--- program cerlatderch (robot Fanuc LR Mate 200iD/7L) ---
  Suave(1)
  Establecer velocidad (1000.0 mm/s)
  Est. Ref.: RobotiQ 2F-140 Gripper (Mechanism) Base
  Est. herr: Tool 1
  Mostrar Tool 1
  MoveJ 1 to (255.53, 172.79, 254.67) mm, rotated rx 167 ry -29.36 rz -83.53 deg; joints [62.819, 42.709, -13.957, -31.792, -82.544, 126.287]
  MoveL 2 to (255.53, 172.79, 254.67) mm, rotated rx 167 ry -29.36 rz -83.53 deg; joints [62.819, 42.709, -13.957, -31.792, -82.544, 126.287]
  MoveL 3 to (235.92, 172.79, 156.61) mm, rotated rx 167 ry -29.36 rz -83.53 deg; joints [63.476, 48.891, -22.926, -32.864, -74.628, 130.64]
  MoveL 4 to (235.92, 172.79, 156.61) mm, rotated rx 167 ry -29.36 rz -83.53 deg; joints [63.476, 48.891, -22.926, -32.864, -74.628, 130.64]
  Establecer velocidad (50.0 mm/s)
  MoveL 5 to (245.19, 173.88, 156.61) mm, rotated rx 167 ry -29.36 rz -83.53 deg; joints [63.097, 47.784, -23.838, -32.935, -74.051, 131.456]
  MoveL 6 to (254.51, 174, 156.61) mm, rotated rx 167 ry -29.36 rz -83.53 deg; joints [62.774, 46.641, -24.767, -33.021, -73.432, 132.241]
  MoveL 7 to (263.84, 173.92, 156.61) mm, rotated rx 167 ry -29.36 rz -83.53 deg; joints [62.457, 45.515, -25.67, -33.109, -72.832, 133.007]
  MoveL 8 to (273.13, 173.41, 156.77) mm, rotated rx 167 ry -29.36 rz -83.53 deg; joints [62.163, 44.386, -26.542, -33.199, -72.246, 133.739]
  MoveL 9 to (282.79, 172.36, 157.79) mm, rotated rx 167 ry -29.36 rz -83.53 deg; joints [61.885, 43.161, -27.346, -33.284, -71.709, 134.42]
  MoveL 10 to (292.21, 170.83, 159.74) mm, rotated rx 167 ry -29.36 rz -83.53 deg; joints [61.643, 41.908, -28.02, -33.355, -71.264, 134.999]
  MoveL 11 to (301.4, 168.84, 162.6) mm, rotated rx 167 ry -29.36 rz -83.53 deg; joints [61.436, 40.621, -28.563, -33.411, -70.911, 135.476]
  MoveL 12 to (310.49, 166.4, 165.63) mm, rotated rx 167 ry -29.36 rz -83.53 deg; joints [61.259, 39.322, -29.065, -33.468, -70.577, 135.906]
  MoveL 13 to (319.81, 164.14, 167.77) mm, rotated rx 167 ry -29.36 rz -83.53 deg; joints [61.056, 38.072, -29.642, -33.535, -70.194, 136.401]
  MoveL 14 to (329.36, 162.38, 169) mm, rotated rx 167 ry -29.36 rz -83.53 deg; joints [60.801, 36.892, -30.285, -33.604, -69.78, 136.975]
  MoveL 15 to (339.84, 161.1, 169.31) mm, rotated rx 167 ry -29.36 rz -83.53 deg; joints [60.468, 35.712, -31.049, -33.681, -69.303, 137.681]
  MoveL 16 to (350.39, 160.46, 169.31) mm, rotated rx 167 ry -29.36 rz -83.53 deg; joints [60.074, 34.597, -31.799, -33.741, -68.866, 138.426]
  MoveL 17 to (360.96, 160.39, 169.31) mm, rotated rx 167 ry -29.36 rz -83.53 deg; joints [59.626, 33.529, -32.502, -33.778, -68.492, 139.185]
  MoveL 18 to (371.53, 160.39, 169.31) mm, rotated rx 167 ry -29.36 rz -83.53 deg; joints [59.16, 32.48, -33.179, -33.805, -68.148, 139.94]
  MoveL 19 to (382.1, 160.39, 169.31) mm, rotated rx 167 ry -29.36 rz -83.53 deg; joints [58.681, 31.444, -33.831, -33.821, -67.828, 140.689]
  MoveL 20 to (408.52, 160.39, 169.31) mm, rotated rx 167 ry -29.36 rz -83.53 deg; joints [57.423, 28.911, -35.364, -33.817, -67.131, 142.544]
  MoveL 21 to (413.03, 160.03, 169.31) mm, rotated rx 167 ry -29.36 rz -83.53 deg; joints [57.227, 28.464, -35.624, -33.821, -67.004, 142.845]
  MoveL 22 to (417.64, 158.65, 169.31) mm, rotated rx 167 ry -29.36 rz -83.53 deg; joints [57.103, 27.947, -35.922, -33.855, -66.812, 143.116]
  MoveL 23 to (422.01, 156.15, 169.31) mm, rotated rx 167 ry -29.36 rz -83.53 deg; joints [57.077, 27.387, -36.239, -33.923, -66.56, 143.328]
  MoveL 24 to (425.74, 152.66, 169.31) mm, rotated rx 167 ry -29.36 rz -83.53 deg; joints [57.162, 26.828, -36.552, -34.025, -66.262, 143.456]
  MoveL 25 to (428.54, 148.44, 169.31) mm, rotated rx 167 ry -29.36 rz -83.53 deg; joints [57.356, 26.314, -36.835, -34.154, -65.941, 143.489]
  MoveL 26 to (430.23, 143.87, 169.31) mm, rotated rx 167 ry -29.36 rz -83.53 deg; joints [57.636, 25.883, -37.068, -34.299, -65.622, 143.43]
  MoveL 27 to (430.87, 139.33, 169.31) mm, rotated rx 167 ry -29.36 rz -83.53 deg; joints [57.973, 25.556, -37.244, -34.446, -65.326, 143.295]
  MoveL 28 to (430.88, 134.93, 169.31) mm, rotated rx 167 ry -29.36 rz -83.53 deg; joints [58.333, 25.298, -37.381, -34.591, -65.05, 143.121]
  MoveL 29 to (430.86, 130.52, 169.31) mm, rotated rx 167 ry -29.36 rz -83.53 deg; joints [58.698, 25.045, -37.514, -34.737, -64.776, 142.942]
  MoveL 30 to (430.2, 125.97, 169.31) mm, rotated rx 167 ry -29.36 rz -83.53 deg; joints [59.109, 24.848, -37.618, -34.889, -64.505, 142.711]
  MoveL 31 to (428.47, 121.41, 169.31) mm, rotated rx 167 ry -29.36 rz -83.53 deg; joints [59.577, 24.755, -37.666, -35.042, -64.253, 142.405]
  MoveL 32 to (425.65, 117.21, 169.31) mm, rotated rx 167 ry -29.36 rz -83.53 deg; joints [60.069, 24.791, -37.647, -35.183, -64.045, 142.039]
  MoveL 33 to (421.9, 113.74, 169.31) mm, rotated rx 167 ry -29.36 rz -83.53 deg; joints [60.543, 24.962, -37.558, -35.297, -63.901, 141.64]
  MoveL 34 to (417.52, 111.28, 169.31) mm, rotated rx 167 ry -29.36 rz -83.53 deg; joints [60.959, 25.251, -37.405, -35.375, -63.834, 141.242]
  MoveL 35 to (412.24, 109.81, 169.31) mm, rotated rx 167 ry -29.36 rz -83.53 deg; joints [61.327, 25.684, -37.175, -35.415, -63.852, 140.827]
  MoveL 36 to (407.14, 109.59, 169.31) mm, rotated rx 167 ry -29.36 rz -83.53 deg; joints [61.58, 26.169, -36.913, -35.413, -63.949, 140.475]
  MoveL 37 to (402.11, 109.59, 169.31) mm, rotated rx 167 ry -29.36 rz -83.53 deg; joints [61.806, 26.66, -36.644, -35.4, -64.063, 140.137]
  MoveL 38 to (397.07, 109.59, 169.31) mm, rotated rx 167 ry -29.36 rz -83.53 deg; joints [62.03, 27.154, -36.37, -35.385, -64.183, 139.798]
  MoveL 39 to (392.04, 109.59, 169.31) mm, rotated rx 167 ry -29.36 rz -83.53 deg; joints [62.25, 27.65, -36.091, -35.367, -64.308, 139.458]
  MoveL 40 to (387.01, 109.59, 169.31) mm, rotated rx 167 ry -29.36 rz -83.53 deg; joints [62.467, 28.147, -35.807, -35.347, -64.438, 139.117]
  MoveL 41 to (381.98, 109.59, 169.31) mm, rotated rx 167 ry -29.36 rz -83.53 deg; joints [62.681, 28.647, -35.517, -35.325, -64.573, 138.774]
  MoveL 42 to (370.35, 109.59, 169.31) mm, rotated rx 167 ry -29.36 rz -83.53 deg; joints [63.163, 29.81, -34.83, -35.263, -64.906, 137.979]
  MoveL 43 to (358.72, 109.59, 169.31) mm, rotated rx 167 ry -29.36 rz -83.53 deg; joints [63.63, 30.986, -34.115, -35.19, -65.268, 137.178]
  MoveL 44 to (347.1, 109.76, 169.31) mm, rotated rx 167 ry -29.36 rz -83.53 deg; joints [64.069, 32.184, -33.366, -35.101, -65.671, 136.376]
  MoveL 45 to (335.47, 109.5, 169.3) mm, rotated rx 167 ry -29.36 rz -83.53 deg; joints [64.527, 33.378, -32.602, -35.013, -66.075, 135.551]
  MoveL 46 to (325.71, 108.73, 168.64) mm, rotated rx 167 ry -29.36 rz -83.53 deg; joints [64.943, 34.406, -32.028, -34.963, -66.344, 134.876]
  MoveL 47 to (316.17, 107.5, 167.04) mm, rotated rx 167 ry -29.36 rz -83.53 deg; joints [65.376, 35.455, -31.568, -34.945, -66.51, 134.259]
  MoveL 48 to (306.86, 105.82, 164.53) mm, rotated rx 167 ry -29.36 rz -83.53 deg; joints [65.826, 36.522, -31.218, -34.955, -66.577, 133.698]
  MoveL 49 to (297.74, 103.7, 161.34) mm, rotated rx 167 ry -29.36 rz -83.53 deg; joints [66.291, 37.598, -30.947, -34.987, -66.571, 133.172]
  MoveL 50 to (288.57, 101.1, 158.87) mm, rotated rx 167 ry -29.36 rz -83.53 deg; joints [66.786, 38.625, -30.584, -34.999, -66.625, 132.566]
  MoveL 51 to (279.32, 97.99, 157.31) mm, rotated rx 167 ry -29.36 rz -83.53 deg; joints [67.309, 39.597, -30.108, -34.986, -66.755, 131.867]
  MoveL 52 to (269.16, 95.14, 156.63) mm, rotated rx 167 ry -29.36 rz -83.53 deg; joints [67.83, 40.652, -29.429, -34.921, -67.053, 131.04]
  MoveL 53 to (258.73, 93.27, 156.61) mm, rotated rx 167 ry -29.36 rz -83.53 deg; joints [68.276, 41.767, -28.59, -34.803, -67.518, 130.173]
  MoveL 54 to (248.13, 92.41, 156.61) mm, rotated rx 167 ry -29.36 rz -83.53 deg; joints [68.643, 42.973, -27.665, -34.652, -68.094, 129.318]
  MoveL 55 to (237.5, 92.57, 156.61) mm, rotated rx 167 ry -29.36 rz -83.53 deg; joints [68.927, 44.261, -26.662, -34.475, -68.777, 128.482]
  MoveL 56 to (226.98, 93.76, 156.67) mm, rotated rx 167 ry -29.36 rz -83.53 deg; joints [69.129, 45.614, -25.583, -34.275, -69.565, 127.669]
  MoveL 57 to (220.53, 95, 156.94) mm, rotated rx 167 ry -29.36 rz -83.53 deg; joints [69.214, 46.476, -24.851, -34.137, -70.127, 127.164]
  MoveL 58 to (214.18, 96.62, 157.45) mm, rotated rx 167 ry -29.36 rz -83.53 deg; joints [69.269, 47.348, -24.072, -33.99, -70.745, 126.656]
  MoveL 59 to (207.94, 98.62, 158.18) mm, rotated rx 167 ry -29.36 rz -83.53 deg; joints [69.294, 48.235, -23.243, -33.835, -71.42, 126.147]
  MoveL 60 to (202.03, 101.35, 159.07) mm, rotated rx 167 ry -29.36 rz -83.53 deg; joints [69.26, 49.127, -22.379, -33.672, -72.155, 125.67]
  MoveL 61 to (196.78, 105.2, 160.04) mm, rotated rx 167 ry -29.36 rz -83.53 deg; joints [69.133, 50.007, -21.509, -33.504, -72.945, 125.267]
  MoveL 62 to (192.41, 110, 160.98) mm, rotated rx 167 ry -29.36 rz -83.53 deg; joints [68.923, 50.84, -20.677, -33.341, -73.747, 124.96]
  MoveL 63 to (189.05, 115.61, 161.78) mm, rotated rx 167 ry -29.36 rz -83.53 deg; joints [68.635, 51.604, -19.92, -33.187, -74.529, 124.763]
  MoveL 64 to (186.87, 121.77, 162.34) mm, rotated rx 167 ry -29.36 rz -83.53 deg; joints [68.284, 52.257, -19.287, -33.05, -75.24, 124.692]
  MoveL 65 to (186.12, 126.11, 162.54) mm, rotated rx 167 ry -29.36 rz -83.53 deg; joints [68.018, 52.62, -18.948, -32.97, -75.661, 124.719]
  MoveL 66 to (185.93, 130.52, 162.58) mm, rotated rx 167 ry -29.36 rz -83.53 deg; joints [67.733, 52.914, -18.69, -32.9, -76.024, 124.807]
  MoveL 67 to (186.01, 134.94, 162.56) mm, rotated rx 167 ry -29.36 rz -83.53 deg; joints [67.443, 53.178, -18.465, -32.834, -76.362, 124.92]
  MoveL 68 to (186.83, 139.23, 162.35) mm, rotated rx 167 ry -29.36 rz -83.53 deg; joints [67.141, 53.335, -18.361, -32.783, -76.605, 125.109]
  MoveL 69 to (189.27, 144.53, 161.73) mm, rotated rx 167 ry -29.36 rz -83.53 deg; joints [66.73, 53.332, -18.45, -32.742, -76.741, 125.496]
  MoveL 70 to (192.92, 149.04, 160.87) mm, rotated rx 167 ry -29.36 rz -83.53 deg; joints [66.335, 53.113, -18.76, -32.73, -76.683, 125.992]
  MoveL 71 to (196.97, 153.16, 160.01) mm, rotated rx 167 ry -29.36 rz -83.53 deg; joints [65.952, 52.817, -19.134, -32.727, -76.564, 126.513]
  MoveL 72 to (203.59, 158.73, 158.82) mm, rotated rx 167 ry -29.36 rz -83.53 deg; joints [65.398, 52.27, -19.77, -32.731, -76.311, 127.319]
  MoveL 73 to (210.87, 163.56, 157.81) mm, rotated rx 167 ry -29.36 rz -83.53 deg; joints [64.867, 51.598, -20.485, -32.747, -75.979, 128.149]
  MoveL 74 to (218.67, 167.53, 157.07) mm, rotated rx 167 ry -29.36 rz -83.53 deg; joints [64.37, 50.814, -21.254, -32.774, -75.585, 128.981]
  MoveL 75 to (226.86, 170.59, 156.67) mm, rotated rx 167 ry -29.36 rz -83.53 deg; joints [63.913, 49.93, -22.054, -32.812, -75.142, 129.798]
  Establecer velocidad (1000.0 mm/s)
  MoveL 76 to (226.86, 170.59, 156.67) mm, rotated rx 167 ry -29.36 rz -83.53 deg; joints [63.913, 49.93, -22.054, -32.812, -75.142, 129.798]
  MoveL 77 to (246.47, 170.59, 254.73) mm, rotated rx 167 ry -29.36 rz -83.53 deg; joints [63.272, 43.813, -13.15, -31.797, -82.998, 125.482]
  Establecer velocidad (1000.0 mm/s)
  MoveL 78 to (401.83, 160.52, 306.49) mm, rotated rx 167 ry -29.36 rz -83.53 deg; joints [57.739, 22.896, -18.143, -31.275, -81.532, 132.699]
  MoveL 79 to (382.22, 160.52, 208.44) mm, rotated rx 167 ry -29.36 rz -83.53 deg; joints [58.665, 29.141, -29.231, -32.884, -71.679, 138.006]
  MoveL 80 to (382.22, 160.52, 208.44) mm, rotated rx 167 ry -29.36 rz -83.53 deg; joints [58.665, 29.141, -29.231, -32.884, -71.679, 138.006]
  Establecer velocidad (50.0 mm/s)
  MoveL 81 to (398.1, 159.77, 208.44) mm, rotated rx 167 ry -29.36 rz -83.53 deg; joints [57.977, 27.495, -30.13, -32.875, -71.248, 139.05]
  MoveL 82 to (413.85, 157.57, 208.44) mm, rotated rx 167 ry -29.36 rz -83.53 deg; joints [57.377, 25.796, -31.013, -32.884, -70.787, 140.016]
  MoveL 83 to (418.98, 156.18, 208.44) mm, rotated rx 167 ry -29.36 rz -83.53 deg; joints [57.228, 25.206, -31.31, -32.901, -70.607, 140.3]
  MoveL 84 to (423.65, 153.71, 208.44) mm, rotated rx 167 ry -29.36 rz -83.53 deg; joints [57.186, 24.593, -31.611, -32.947, -70.373, 140.506]
  MoveL 85 to (427.7, 150.29, 208.44) mm, rotated rx 167 ry -29.36 rz -83.53 deg; joints [57.25, 23.982, -31.906, -33.022, -70.097, 140.627]
  MoveL 86 to (430.9, 146.07, 208.44) mm, rotated rx 167 ry -29.36 rz -83.53 deg; joints [57.424, 23.406, -32.178, -33.124, -69.788, 140.654]
  MoveL 87 to (432.92, 141.18, 208.44) mm, rotated rx 167 ry -29.36 rz -83.53 deg; joints [57.717, 22.905, -32.409, -33.25, -69.459, 140.568]
  MoveL 88 to (433.51, 135.92, 208.44) mm, rotated rx 167 ry -29.36 rz -83.53 deg; joints [58.117, 22.524, -32.583, -33.395, -69.128, 140.369]
  MoveL 89 to (433.26, 130.66, 208.44) mm, rotated rx 167 ry -29.36 rz -83.53 deg; joints [58.565, 22.229, -32.715, -33.544, -68.81, 140.11]
  MoveL 90 to (431.75, 125.64, 208.44) mm, rotated rx 167 ry -29.36 rz -83.53 deg; joints [59.059, 22.078, -32.783, -33.69, -68.524, 139.778]
  MoveL 91 to (428.97, 121.16, 208.44) mm, rotated rx 167 ry -29.36 rz -83.53 deg; joints [59.573, 22.09, -32.777, -33.825, -68.288, 139.389]
  MoveL 92 to (425.29, 117.41, 208.44) mm, rotated rx 167 ry -29.36 rz -83.53 deg; joints [60.069, 22.241, -32.71, -33.94, -68.111, 138.975]
  MoveL 93 to (421.02, 114.59, 208.44) mm, rotated rx 167 ry -29.36 rz -83.53 deg; joints [60.513, 22.508, -32.59, -34.027, -68.002, 138.569]
  MoveL 94 to (416.24, 112.78, 208.44) mm, rotated rx 167 ry -29.36 rz -83.53 deg; joints [60.891, 22.888, -32.417, -34.085, -67.967, 138.179]
  MoveL 95 to (411.24, 111.87, 208.44) mm, rotated rx 167 ry -29.36 rz -83.53 deg; joints [61.2, 23.343, -32.206, -34.115, -67.995, 137.819]
  MoveL 96 to (406.21, 111.14, 208.44) mm, rotated rx 167 ry -29.36 rz -83.53 deg; joints [61.491, 23.815, -31.985, -34.137, -68.04, 137.464]
  MoveL 97 to (393.32, 109.92, 208.44) mm, rotated rx 167 ry -29.36 rz -83.53 deg; joints [62.167, 25.068, -31.378, -34.164, -68.22, 136.585]
  MoveL 98 to (380.38, 109.57, 208.44) mm, rotated rx 167 ry -29.36 rz -83.53 deg; joints [62.749, 26.389, -30.71, -34.151, -68.492, 135.737]
  MoveL 99 to (368.61, 109.92, 208.44) mm, rotated rx 167 ry -29.36 rz -83.53 deg; joints [63.207, 27.639, -30.053, -34.111, -68.815, 134.99]
  MoveL 100 to (356.97, 111.21, 208.44) mm, rotated rx 167 ry -29.36 rz -83.53 deg; joints [63.57, 28.939, -29.343, -34.038, -69.225, 134.285]
  MoveL 101 to (345.55, 113.37, 208.44) mm, rotated rx 167 ry -29.36 rz -83.53 deg; joints [63.844, 30.275, -28.588, -33.939, -69.717, 133.622]
  MoveL 102 to (333.92, 113.25, 208.44) mm, rotated rx 167 ry -29.36 rz -83.53 deg; joints [64.293, 31.528, -27.855, -33.881, -70.105, 132.837]
  MoveL 103 to (322.29, 113.18, 208.44) mm, rotated rx 167 ry -29.36 rz -83.53 deg; joints [64.724, 32.803, -27.087, -33.814, -70.53, 132.045]
  MoveL 104 to (318.84, 113.27, 208.44) mm, rotated rx 167 ry -29.36 rz -83.53 deg; joints [64.842, 33.192, -26.849, -33.79, -70.669, 131.812]
  MoveL 105 to (315.38, 113.44, 208.44) mm, rotated rx 167 ry -29.36 rz -83.53 deg; joints [64.952, 33.586, -26.605, -33.763, -70.818, 131.582]
  MoveL 106 to (311.94, 113.73, 208.44) mm, rotated rx 167 ry -29.36 rz -83.53 deg; joints [65.051, 33.988, -26.353, -33.733, -70.977, 131.356]
  MoveL 107 to (308.53, 114.29, 208.44) mm, rotated rx 167 ry -29.36 rz -83.53 deg; joints [65.128, 34.401, -26.093, -33.698, -71.156, 131.142]
  MoveL 108 to (305.51, 115.94, 208.44) mm, rotated rx 167 ry -29.36 rz -83.53 deg; joints [65.11, 34.829, -25.821, -33.644, -71.391, 130.998]
  MoveL 109 to (303.55, 118.04, 208.44) mm, rotated rx 167 ry -29.36 rz -83.53 deg; joints [65.021, 35.163, -25.606, -33.588, -71.614, 130.943]
  MoveL 110 to (302.26, 120.61, 208.44) mm, rotated rx 167 ry -29.36 rz -83.53 deg; joints [64.874, 35.447, -25.423, -33.528, -71.84, 130.952]
  MoveL 111 to (301.89, 123.45, 208.44) mm, rotated rx 167 ry -29.36 rz -83.53 deg; joints [64.677, 35.642, -25.297, -33.469, -72.044, 131.035]
  MoveL 112 to (302.49, 126.27, 208.44) mm, rotated rx 167 ry -29.36 rz -83.53 deg; joints [64.448, 35.726, -25.242, -33.417, -72.204, 131.185]
  MoveL 113 to (303.41, 129.02, 208.44) mm, rotated rx 167 ry -29.36 rz -83.53 deg; joints [64.213, 35.772, -25.213, -33.368, -72.345, 131.354]
  MoveL 114 to (304.36, 131.76, 208.44) mm, rotated rx 167 ry -29.36 rz -83.53 deg; joints [63.978, 35.816, -25.184, -33.32, -72.486, 131.524]
  MoveL 115 to (304.62, 133.96, 208.44) mm, rotated rx 167 ry -29.36 rz -83.53 deg; joints [63.808, 35.909, -25.123, -33.277, -72.621, 131.624]
  MoveL 116 to (303.96, 136.18, 208.44) mm, rotated rx 167 ry -29.36 rz -83.53 deg; joints [63.669, 36.109, -24.993, -33.229, -72.799, 131.659]
  MoveL 117 to (303.31, 138.41, 208.44) mm, rotated rx 167 ry -29.36 rz -83.53 deg; joints [63.531, 36.308, -24.862, -33.181, -72.978, 131.694]
  MoveL 118 to (302.68, 140.64, 208.44) mm, rotated rx 167 ry -29.36 rz -83.53 deg; joints [63.392, 36.507, -24.73, -33.133, -73.157, 131.729]
  MoveL 119 to (302.1, 142.88, 208.44) mm, rotated rx 167 ry -29.36 rz -83.53 deg; joints [63.251, 36.703, -24.601, -33.085, -73.335, 131.767]
  MoveL 120 to (302.05, 146.74, 208.44) mm, rotated rx 167 ry -29.36 rz -83.53 deg; joints [62.975, 36.931, -24.449, -33.008, -73.599, 131.9]
  MoveL 121 to (303.35, 150.38, 208.44) mm, rotated rx 167 ry -29.36 rz -83.53 deg; joints [62.667, 36.996, -24.406, -32.943, -73.788, 132.121]
  MoveL 122 to (305.63, 153.5, 208.44) mm, rotated rx 167 ry -29.36 rz -83.53 deg; joints [62.359, 36.922, -24.455, -32.892, -73.899, 132.394]
  MoveL 123 to (308.22, 155.56, 208.44) mm, rotated rx 167 ry -29.36 rz -83.53 deg; joints [62.114, 36.75, -24.569, -32.862, -73.924, 132.653]
  MoveL 124 to (311.4, 156.56, 208.44) mm, rotated rx 167 ry -29.36 rz -83.53 deg; joints [61.923, 36.452, -24.767, -32.855, -73.852, 132.917]
  MoveL 125 to (314.73, 157, 208.44) mm, rotated rx 167 ry -29.36 rz -83.53 deg; joints [61.763, 36.105, -24.995, -32.859, -73.739, 133.172]
  MoveL 126 to (318.08, 157.27, 208.44) mm, rotated rx 167 ry -29.36 rz -83.53 deg; joints [61.615, 35.747, -25.229, -32.866, -73.616, 133.422]
  MoveL 127 to (321.43, 157.41, 208.44) mm, rotated rx 167 ry -29.36 rz -83.53 deg; joints [61.474, 35.383, -25.465, -32.876, -73.487, 133.667]
  MoveL 128 to (324.78, 157.45, 208.44) mm, rotated rx 167 ry -29.36 rz -83.53 deg; joints [61.34, 35.016, -25.701, -32.886, -73.354, 133.907]
  MoveL 129 to (328.13, 157.42, 208.44) mm, rotated rx 167 ry -29.36 rz -83.53 deg; joints [61.209, 34.647, -25.937, -32.897, -73.22, 134.144]
  MoveL 130 to (335.01, 157.24, 208.44) mm, rotated rx 167 ry -29.36 rz -83.53 deg; joints [60.946, 33.887, -26.417, -32.921, -72.945, 134.624]
  MoveL 131 to (341.89, 157.02, 208.44) mm, rotated rx 167 ry -29.36 rz -83.53 deg; joints [60.681, 33.133, -26.886, -32.942, -72.681, 135.099]
  MoveL 132 to (348.73, 157.41, 208.44) mm, rotated rx 167 ry -29.36 rz -83.53 deg; joints [60.368, 32.427, -27.317, -32.947, -72.47, 135.589]
  MoveL 133 to (355.61, 159.03, 208.44) mm, rotated rx 167 ry -29.36 rz -83.53 deg; joints [59.957, 31.799, -27.695, -32.919, -72.351, 136.126]
  MoveL 134 to (359.78, 159.91, 208.44) mm, rotated rx 167 ry -29.36 rz -83.53 deg; joints [59.712, 31.415, -27.923, -32.902, -72.277, 136.447]
  MoveL 135 to (363.08, 160.33, 208.44) mm, rotated rx 167 ry -29.36 rz -83.53 deg; joints [59.538, 31.096, -28.111, -32.894, -72.203, 136.69]
  MoveL 136 to (365.62, 160.48, 208.44) mm, rotated rx 167 ry -29.36 rz -83.53 deg; joints [59.414, 30.842, -28.26, -32.891, -72.137, 136.871]
  MoveL 137 to (367.82, 160.52, 208.44) mm, rotated rx 167 ry -29.36 rz -83.53 deg; joints [59.315, 30.617, -28.391, -32.891, -72.075, 137.023]
  MoveL 138 to (370.1, 160.52, 208.44) mm, rotated rx 167 ry -29.36 rz -83.53 deg; joints [59.213, 30.381, -28.527, -32.891, -72.009, 137.18]
  MoveL 139 to (372.32, 160.52, 208.44) mm, rotated rx 167 ry -29.36 rz -83.53 deg; joints [59.114, 30.153, -28.659, -32.89, -71.946, 137.332]
  MoveL 140 to (375.19, 160.52, 208.44) mm, rotated rx 167 ry -29.36 rz -83.53 deg; joints [58.985, 29.859, -28.827, -32.889, -71.866, 137.527]
  MoveL 141 to (378.62, 160.52, 208.44) mm, rotated rx 167 ry -29.36 rz -83.53 deg; joints [58.83, 29.508, -29.025, -32.887, -71.773, 137.761]
  MoveL 142 to (382.22, 160.52, 208.44) mm, rotated rx 167 ry -29.36 rz -83.53 deg; joints [58.665, 29.141, -29.231, -32.884, -71.679, 138.006]
  Establecer velocidad (1000.0 mm/s)
  MoveL 143 to (382.22, 160.52, 208.44) mm, rotated rx 167 ry -29.36 rz -83.53 deg; joints [58.665, 29.141, -29.231, -32.884, -71.679, 138.006]
  MoveL 144 to (401.83, 160.52, 306.49) mm, rotated rx 167 ry -29.36 rz -83.53 deg; joints [57.739, 22.896, -18.143, -31.275, -81.532, 132.699]

--- program ceraarribderch (robot Fanuc LR Mate 200iD/7L) ---
  Suave(1)
  Establecer velocidad (1000.0 mm/s)
  Est. Ref.: bote cera
  Est. herr: Tool 1
  Mostrar Tool 1
  MoveJ 1 to (349.44, 103.38, 195.99) mm, rotated rx 122.56 ry -24.48 rz -84.76 deg; joints [61.244, 18.633, -53.476, -104.529, -42.664, -159.742]
  MoveL 2 to (349.44, 103.38, 195.99) mm, rotated rx 122.56 ry -24.48 rz -84.76 deg; joints [61.244, 18.633, -53.476, -104.529, -42.664, -159.742]
  MoveL 3 to (329.83, 103.38, 97.93) mm, rotated rx 122.56 ry -24.48 rz -84.76 deg; joints [62.357, 32.195, -66.199, -117.758, -46.769, -142.563]
  MoveL 4 to (329.83, 103.38, 97.93) mm, rotated rx 122.56 ry -24.48 rz -84.76 deg; joints [62.357, 32.195, -66.199, -117.758, -46.769, -142.563]
  Establecer velocidad (50.0 mm/s)
  MoveL 5 to (328.15, 103.38, 97.77) mm, rotated rx 122.56 ry -24.48 rz -84.76 deg; joints [62.448, 32.321, -66.096, -117.772, -46.689, -142.664]
  MoveL 6 to (326.47, 103.38, 97.62) mm, rotated rx 122.56 ry -24.48 rz -84.76 deg; joints [62.539, 32.448, -65.992, -117.785, -46.608, -142.766]
  MoveL 7 to (322.21, 103.38, 97.19) mm, rotated rx 122.56 ry -24.48 rz -84.76 deg; joints [62.767, 32.775, -65.732, -117.817, -46.404, -143.023]
  MoveL 8 to (312.54, 103.38, 96.02) mm, rotated rx 122.56 ry -24.48 rz -84.76 deg; joints [63.273, 33.544, -65.159, -117.885, -45.95, -143.589]
  MoveL 9 to (290.7, 103.38, 92.42) mm, rotated rx 122.56 ry -24.48 rz -84.76 deg; joints [64.353, 35.413, -63.937, -118.011, -44.967, -144.799]
  MoveL 10 to (282.18, 103.38, 90.65) mm, rotated rx 122.56 ry -24.48 rz -84.76 deg; joints [64.752, 36.19, -63.484, -118.051, -44.599, -145.248]
  MoveL 11 to (277.43, 103.38, 89.57) mm, rotated rx 122.56 ry -24.48 rz -84.76 deg; joints [64.97, 36.634, -63.237, -118.07, -44.396, -145.494]
  MoveL 12 to (274.78, 103.38, 88.94) mm, rotated rx 122.56 ry -24.48 rz -84.76 deg; joints [65.09, 36.886, -63.101, -118.08, -44.284, -145.63]
  MoveL 13 to (273.09, 103.38, 88.53) mm, rotated rx 122.56 ry -24.48 rz -84.76 deg; joints [65.166, 37.048, -63.014, -118.086, -44.213, -145.715]
  MoveL 14 to (271.43, 103.38, 88.06) mm, rotated rx 122.56 ry -24.48 rz -84.76 deg; joints [65.24, 37.215, -62.937, -118.098, -44.147, -145.791]
  MoveL 15 to (269.69, 103.38, 86.4) mm, rotated rx 122.56 ry -24.48 rz -84.76 deg; joints [65.318, 37.526, -62.988, -118.231, -44.14, -145.702]
  MoveL 16 to (269.33, 103.38, 85.24) mm, rotated rx 122.56 ry -24.48 rz -84.76 deg; joints [65.334, 37.688, -63.092, -118.343, -44.183, -145.565]
  MoveL 17 to (269.29, 103.38, 84.03) mm, rotated rx 122.56 ry -24.48 rz -84.76 deg; joints [65.335, 37.834, -63.229, -118.468, -44.247, -145.393]
  MoveL 18 to (269.29, 103.38, 79.16) mm, rotated rx 122.56 ry -24.48 rz -84.76 deg; joints [65.335, 38.413, -63.785, -118.967, -44.515, -144.695]
  MoveL 19 to (269.29, 103.38, 69.43) mm, rotated rx 122.56 ry -24.48 rz -84.76 deg; joints [65.335, 39.581, -64.884, -119.931, -45.055, -143.337]
  Establecer velocidad (1000.0 mm/s)
  MoveL 20 to (269.29, 103.38, 69.43) mm, rotated rx 122.56 ry -24.48 rz -84.76 deg; joints [65.335, 39.581, -64.884, -119.931, -45.055, -143.337]
  MoveL 21 to (288.9, 103.38, 167.49) mm, rotated rx 122.56 ry -24.48 rz -84.76 deg; joints [64.438, 26.897, -54.3, -108.589, -41.095, -157.756]
  Establecer velocidad (1000.0 mm/s)
  MoveL 22 to (349.44, 103.38, 195.99) mm, rotated rx 122.56 ry -24.48 rz -84.76 deg; joints [61.244, 18.633, -53.476, -104.529, -42.664, -159.742]
  MoveL 23 to (329.83, 103.38, 97.93) mm, rotated rx 122.56 ry -24.48 rz -84.76 deg; joints [62.357, 32.195, -66.199, -117.758, -46.769, -142.563]
  MoveL 24 to (329.83, 103.38, 97.93) mm, rotated rx 122.56 ry -24.48 rz -84.76 deg; joints [62.357, 32.195, -66.199, -117.758, -46.769, -142.563]
  Establecer velocidad (50.0 mm/s)
  MoveL 25 to (342.28, 103.38, 99.54) mm, rotated rx 122.56 ry -24.48 rz -84.76 deg; joints [61.66, 31.199, -66.891, -117.57, -47.336, -141.9]
  MoveL 26 to (354.55, 103.38, 102.17) mm, rotated rx 122.56 ry -24.48 rz -84.76 deg; joints [60.941, 30.078, -67.406, -117.208, -47.821, -141.454]
  MoveL 27 to (366.58, 103.38, 105.81) mm, rotated rx 122.56 ry -24.48 rz -84.76 deg; joints [60.204, 28.827, -67.729, -116.67, -48.218, -141.24]
  MoveL 28 to (378.26, 103.38, 110.44) mm, rotated rx 122.56 ry -24.48 rz -84.76 deg; joints [59.454, 27.444, -67.842, -115.955, -48.522, -141.272]
  MoveL 29 to (392.5, 103.38, 117.7) mm, rotated rx 122.56 ry -24.48 rz -84.76 deg; joints [58.493, 25.497, -67.662, -114.785, -48.774, -141.696]
  MoveL 30 to (405.91, 103.38, 126.43) mm, rotated rx 122.56 ry -24.48 rz -84.76 deg; joints [57.537, 23.347, -67.102, -113.324, -48.881, -142.575]
  MoveL 31 to (418.33, 103.38, 136.51) mm, rotated rx 122.56 ry -24.48 rz -84.76 deg; joints [56.605, 21.011, -66.148, -111.575, -48.859, -143.933]
  MoveL 32 to (429.62, 103.38, 147.83) mm, rotated rx 122.56 ry -24.48 rz -84.76 deg; joints [55.715, 18.518, -64.801, -109.548, -48.732, -145.781]
  Establecer velocidad (1000.0 mm/s)
  MoveL 33 to (429.62, 103.38, 147.83) mm, rotated rx 122.56 ry -24.48 rz -84.76 deg; joints [55.715, 18.518, -64.801, -109.548, -48.732, -145.781]
  MoveL 34 to (449.23, 103.38, 245.88) mm, rotated rx 122.56 ry -24.48 rz -84.76 deg; joints [54.067, 3.573, -48.055, -92.811, -46.344, -168.354]
  Establecer velocidad (1000.0 mm/s)
  MoveL 35 to (530.22, 103.38, 245.88) mm, rotated rx 122.56 ry -24.48 rz -84.76 deg; joints [45.585, -4.583, -47.952, -86.445, -52.017, -168.441]
  MoveL 36 to (510.6, 103.38, 147.83) mm, rotated rx 122.56 ry -24.48 rz -84.76 deg; joints [47.924, 12.844, -68.18, -104.299, -52.686, -142.783]
  MoveL 37 to (510.6, 103.38, 147.83) mm, rotated rx 122.56 ry -24.48 rz -84.76 deg; joints [47.924, 12.844, -68.18, -104.299, -52.686, -142.783]
  Establecer velocidad (50.0 mm/s)
  MoveL 38 to (512.43, 103.38, 137.3) mm, rotated rx 122.56 ry -24.48 rz -84.76 deg; joints [47.715, 14.681, -70.447, -105.738, -53.345, -140.066]
  MoveL 39 to (514.48, 103.38, 126.83) mm, rotated rx 122.56 ry -24.48 rz -84.76 deg; joints [47.478, 16.56, -72.725, -107.104, -54.061, -137.38]
  MoveL 40 to (516.62, 103.38, 116.36) mm, rotated rx 122.56 ry -24.48 rz -84.76 deg; joints [47.229, 18.49, -75.011, -108.405, -54.824, -134.73]
  MoveL 41 to (517.73, 103.38, 106.23) mm, rotated rx 122.56 ry -24.48 rz -84.76 deg; joints [47.098, 20.458, -77.173, -109.692, -55.56, -132.253]
  MoveL 42 to (517.7, 103.38, 96.06) mm, rotated rx 122.56 ry -24.48 rz -84.76 deg; joints [47.102, 22.52, -79.26, -111.02, -56.285, -129.891]
  MoveL 43 to (516.53, 103.38, 86.03) mm, rotated rx 122.56 ry -24.48 rz -84.76 deg; joints [47.239, 24.616, -81.211, -112.355, -56.984, -127.71]
  MoveL 44 to (514.23, 103.38, 76.16) mm, rotated rx 122.56 ry -24.48 rz -84.76 deg; joints [47.507, 26.716, -83.001, -113.687, -57.651, -125.735]
  Establecer velocidad (1000.0 mm/s)
  MoveL 45 to (514.23, 103.38, 76.16) mm, rotated rx 122.56 ry -24.48 rz -84.76 deg; joints [47.507, 26.716, -83.001, -113.687, -57.651, -125.735]
  MoveL 46 to (533.85, 103.38, 174.22) mm, rotated rx 122.56 ry -24.48 rz -84.76 deg; joints [45.131, 6.329, -63.131, -97.816, -52.848, -149.284]

--- program ceraarribaizqch (robot Fanuc LR Mate 200iD/7L) ---
  Suave(1)
  Establecer velocidad (1000.0 mm/s)
  Est. Ref.: RobotiQ 2F-140 Gripper (Mechanism) Base
  Est. herr: Tool 1
  Mostrar Tool 1
  MoveJ 1 to (235.6, -30.8, 267.73) mm, rotated rx 167.98 ry -19.59 rz -85.91 deg; joints [81.108, 34.584, -14.834, -23.134, -68.852, 108.138]
  MoveL 2 to (235.6, -30.8, 267.73) mm, rotated rx 167.98 ry -19.59 rz -85.91 deg; joints [81.108, 34.584, -14.834, -23.134, -68.852, 108.138]
  MoveL 3 to (215.99, -30.8, 169.67) mm, rotated rx 167.98 ry -19.59 rz -85.91 deg; joints [81.345, 40.798, -24.539, -25.02, -59.896, 112.299]
  MoveL 4 to (215.99, -30.8, 169.67) mm, rotated rx 167.98 ry -19.59 rz -85.91 deg; joints [81.345, 40.798, -24.539, -25.02, -59.896, 112.299]
  Establecer velocidad (50.0 mm/s)
  MoveL 5 to (208.21, -30.8, 168.75) mm, rotated rx 167.98 ry -19.59 rz -85.91 deg; joints [81.435, 41.859, -23.896, -24.859, -60.444, 111.9]
  MoveL 6 to (200.43, -30.8, 167.66) mm, rotated rx 167.98 ry -19.59 rz -85.91 deg; joints [81.524, 42.944, -23.245, -24.7, -61.001, 111.503]
  MoveL 7 to (191.82, -30.8, 166.26) mm, rotated rx 167.98 ry -19.59 rz -85.91 deg; joints [81.62, 44.174, -22.514, -24.527, -61.628, 111.065]
  MoveL 8 to (182.09, -30.8, 164.43) mm, rotated rx 167.98 ry -19.59 rz -85.91 deg; joints [81.725, 45.603, -21.672, -24.334, -62.355, 110.569]
  MoveL 9 to (173.76, -30.8, 162.65) mm, rotated rx 167.98 ry -19.59 rz -85.91 deg; joints [81.814, 46.864, -20.933, -24.17, -62.995, 110.143]
  MoveL 10 to (169.82, -30.8, 161.74) mm, rotated rx 167.98 ry -19.59 rz -85.91 deg; joints [81.855, 47.474, -20.576, -24.093, -63.305, 109.94]
  MoveL 11 to (166.31, -30.8, 160.89) mm, rotated rx 167.98 ry -19.59 rz -85.91 deg; joints [81.891, 48.022, -20.256, -24.025, -63.583, 109.759]
  MoveL 12 to (164.84, -30.8, 160.46) mm, rotated rx 167.98 ry -19.59 rz -85.91 deg; joints [81.906, 48.257, -20.127, -23.998, -63.695, 109.686]
  MoveL 13 to (163.89, -30.8, 159.84) mm, rotated rx 167.98 ry -19.59 rz -85.91 deg; joints [81.916, 48.423, -20.08, -23.988, -63.735, 109.656]
  MoveL 14 to (163.09, -30.8, 158.79) mm, rotated rx 167.98 ry -19.59 rz -85.91 deg; joints [81.924, 48.586, -20.096, -23.99, -63.717, 109.655]
  MoveL 15 to (162.75, -30.8, 157.79) mm, rotated rx 167.98 ry -19.59 rz -85.91 deg; joints [81.928, 48.678, -20.162, -24.003, -63.655, 109.682]
  MoveL 16 to (162.68, -30.8, 156.57) mm, rotated rx 167.98 ry -19.59 rz -85.91 deg; joints [81.928, 48.738, -20.286, -24.028, -63.542, 109.737]
  MoveL 17 to (162.68, -30.8, 154.91) mm, rotated rx 167.98 ry -19.59 rz -85.91 deg; joints [81.928, 48.808, -20.463, -24.064, -63.38, 109.818]
  MoveL 18 to (162.68, -30.8, 151.97) mm, rotated rx 167.98 ry -19.59 rz -85.91 deg; joints [81.928, 48.932, -20.776, -24.129, -63.094, 109.961]
  MoveL 19 to (162.68, -30.8, 148.56) mm, rotated rx 167.98 ry -19.59 rz -85.91 deg; joints [81.928, 49.079, -21.138, -24.204, -62.764, 110.128]
  MoveL 20 to (162.68, -30.8, 145.15) mm, rotated rx 167.98 ry -19.59 rz -85.91 deg; joints [81.928, 49.23, -21.499, -24.281, -62.435, 110.294]
  MoveL 21 to (162.68, -30.8, 141.65) mm, rotated rx 167.98 ry -19.59 rz -85.91 deg; joints [81.928, 49.387, -21.866, -24.361, -62.1, 110.466]
  Establecer velocidad (1000.0 mm/s)
  MoveL 22 to (162.68, -30.8, 141.65) mm, rotated rx 167.98 ry -19.59 rz -85.91 deg; joints [81.928, 49.387, -21.866, -24.361, -62.1, 110.466]
  MoveL 23 to (182.3, -30.8, 239.7) mm, rotated rx 167.98 ry -19.59 rz -85.91 deg; joints [81.723, 43.057, -13.081, -22.822, -70.233, 106.822]
  Establecer velocidad (1000.0 mm/s)
  MoveL 24 to (243.44, -30.8, 268.49) mm, rotated rx 167.98 ry -19.59 rz -85.91 deg; joints [81.01, 33.481, -15.383, -23.227, -68.384, 108.464]
  MoveL 25 to (223.83, -30.8, 170.43) mm, rotated rx 167.98 ry -19.59 rz -85.91 deg; joints [81.252, 39.752, -25.18, -25.185, -59.351, 112.703]
  MoveL 26 to (223.83, -30.8, 170.43) mm, rotated rx 167.98 ry -19.59 rz -85.91 deg; joints [81.252, 39.752, -25.18, -25.185, -59.351, 112.703]
  Establecer velocidad (50.0 mm/s)
  MoveL 27 to (238.63, -30.8, 172.45) mm, rotated rx 167.98 ry -19.59 rz -85.91 deg; joints [81.071, 37.785, -26.264, -25.475, -58.441, 113.416]
  MoveL 28 to (254.89, -30.8, 176.41) mm, rotated rx 167.98 ry -19.59 rz -85.91 deg; joints [80.863, 35.58, -27.166, -25.729, -57.708, 114.073]
  MoveL 29 to (270.62, -30.8, 182.12) mm, rotated rx 167.98 ry -19.59 rz -85.91 deg; joints [80.653, 33.381, -27.733, -25.896, -57.279, 114.565]
  MoveL 30 to (285.63, -30.8, 189.51) mm, rotated rx 167.98 ry -19.59 rz -85.91 deg; joints [80.443, 31.202, -27.961, -25.97, -57.154, 114.882]
  MoveL 31 to (299.75, -30.8, 198.51) mm, rotated rx 167.98 ry -19.59 rz -85.91 deg; joints [80.237, 29.059, -27.853, -25.949, -57.332, 115.02]
  MoveL 32 to (312.79, -30.8, 208.99) mm, rotated rx 167.98 ry -19.59 rz -85.91 deg; joints [80.039, 26.978, -27.414, -25.835, -57.803, 114.98]
  MoveL 33 to (324.62, -30.8, 220.83) mm, rotated rx 167.98 ry -19.59 rz -85.91 deg; joints [79.852, 24.986, -26.658, -25.64, -58.556, 114.771]
  Establecer velocidad (1000.0 mm/s)
  MoveL 34 to (324.62, -30.8, 220.83) mm, rotated rx 167.98 ry -19.59 rz -85.91 deg; joints [79.852, 24.986, -26.658, -25.64, -58.556, 114.771]
  MoveL 35 to (344.23, -30.8, 318.89) mm, rotated rx 167.98 ry -19.59 rz -85.91 deg; joints [79.526, 18.985, -15.201, -23.319, -69.117, 109.797]
  Establecer velocidad (1000.0 mm/s)
  MoveL 36 to (426.02, -30.8, 318.89) mm, rotated rx 167.98 ry -19.59 rz -85.91 deg; joints [77.912, 8.736, -17.816, -23.845, -67.34, 112.451]
  MoveL 37 to (406.41, -30.8, 220.83) mm, rotated rx 167.98 ry -19.59 rz -85.91 deg; joints [78.343, 15.384, -30.435, -26.763, -55.752, 118.171]
  MoveL 38 to (406.41, -30.8, 220.83) mm, rotated rx 167.98 ry -19.59 rz -85.91 deg; joints [78.343, 15.384, -30.435, -26.763, -55.752, 118.171]
  Establecer velocidad (50.0 mm/s)
  MoveL 39 to (411.65, -30.8, 193.34) mm, rotated rx 167.98 ry -19.59 rz -85.91 deg; joints [78.231, 16.474, -34.3, -28.055, -52.364, 120.472]
  MoveL 40 to (411.65, -30.8, 193.34) mm, rotated rx 167.98 ry -19.59 rz -85.91 deg; joints [78.231, 16.474, -34.3, -28.055, -52.364, 120.472]
  MoveL 41 to (413.5, -30.8, 180.59) mm, rotated rx 167.98 ry -19.59 rz -85.91 deg; joints [78.191, 17.129, -36.08, -28.726, -50.813, 121.589]
  MoveL 42 to (413.53, -30.8, 167.72) mm, rotated rx 167.98 ry -19.59 rz -85.91 deg; joints [78.191, 18.049, -37.806, -29.428, -49.305, 122.684]
  MoveL 43 to (411.73, -30.8, 154.96) mm, rotated rx 167.98 ry -19.59 rz -85.91 deg; joints [78.23, 19.205, -39.43, -30.141, -47.881, 123.724]
  MoveL 44 to (410.08, -30.8, 148.44) mm, rotated rx 167.98 ry -19.59 rz -85.91 deg; joints [78.265, 19.89, -40.22, -30.507, -47.184, 124.233]
  Establecer velocidad (1000.0 mm/s)
  MoveL 45 to (410.08, -30.8, 148.44) mm, rotated rx 167.98 ry -19.59 rz -85.91 deg; joints [78.265, 19.89, -40.22, -30.507, -47.184, 124.233]
  MoveL 46 to (429.69, -30.8, 246.5) mm, rotated rx 167.98 ry -19.59 rz -85.91 deg; joints [77.829, 11.228, -27.7, -25.988, -58.402, 117.204]

--- program final_ch (robot Fanuc LR Mate 200iD/7L) ---
  Llamar home
  Llamar reset
  Llamar c1 recoger
  Llamar poscharolamesa
  Llamar home
  Llamar iman izquierdo
  Llamar iman derecho
  Llamar recoger cepillo limpi...: recoger cepillo limpieza
  Llamar platizch
  Llamar arrizch
  Llamar pladerch
  Llamar arriderch
  Llamar dejar cepillo limpieza
  Llamar recoger cera
  Llamar cerlatizqch
  Llamar ceraarribaizqch
  Llamar cerlatderch
  Llamar ceraarribderch
  Llamar dejar  cera
  Llamar recoger cepillo cera
  Llamar platizch
  Llamar pladerch
  Llamar arriderch
  Llamar arrizch
  Llamar dejar cepillo cera
  Llamar dejar iman izquierdo
  Llamar home
  Llamar dejar iman derecho
  Llamar pick charola
  Llamar c1 entregar

--- program final_gr (robot Fanuc LR Mate 200iD/7L) ---
  Llamar home
  Llamar reset
  Llamar c1 recoger
  Llamar poscharolamesa
  Llamar home
  Llamar iman izquierdo
  Llamar iman derecho
  Llamar recoger cepillo limpi...: recoger cepillo limpieza
  Llamar plaizgr
  Llamar arriizqgr
  Llamar pladergr
  Llamar arridergr
  Llamar dejar cepillo limpieza
  Llamar recoger cera
  Llamar cerlaizgr
  Llamar ceraariizgr
  Llamar cerladergr
  Llamar cerarridergr
  Llamar dejar  cera
  Llamar recoger cepillo cera
  Llamar plaizgr
  Llamar pladergr
  Llamar arriizqgr
  Llamar arridergr
  Llamar dejar cepillo cera
  Llamar dejar iman izquierdo
  Llamar home
  Llamar dejar iman derecho
  Llamar pick charola
  Llamar c1 entregar
